{attribute 'qualified_only'}
{attribute 'strict'}
TYPE E_HeatPumpAirControlMode :
(
	heatingMode := 2, 
	coolingMode := 3
);
END_TYPE

(* stored: Version 1.1.0.1
   DUT E_HeatPumpAirControlMode: Id {e9df4f15-d1f0-401d-8316-54c8e91f2bd2} *)
